Fanuc KAREL source: kd00031.KL

-- PROVISIONAL review KL for V940-1; original PC SHA256 3eebfd0d5bb816f11aa05a0620538a37a3ce10d994448d58d85b1018d59421e1
-- Incomplete behavior may be omitted. Consult companion uncertainty JSON. Do not deploy.
PROGRAM KD00031
%NOLOCKGROUP
VAR
  I : INTEGER
  J : INTEGER
  B : BOOLEAN
  R : REAL
  S : STRING[80]
BEGIN
  -- V9_ZERO_TABLE_METADATA_HINT layout=0001; no indexed target words; source/name/runtime held
  -- UNRESOLVED_PC offsets 5-21; opcodes 9D,81,18,9C,12,22,9D,13,04
  -- UNRESOLVED_PC offsets 26-30; opcodes 7F
END KD00031
